// TIA Portal V21 export
ORGANIZATION_BLOCK "Pair"   // OB1, LAD
BEGIN

REGION Network 1: Motor
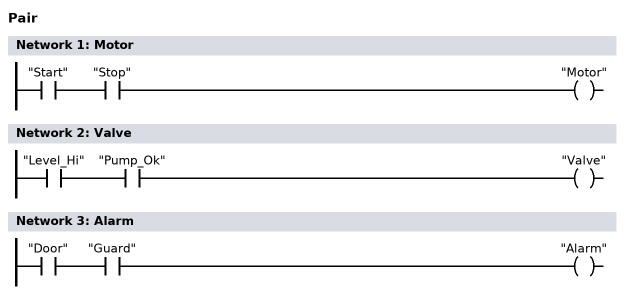
   RUNG wire#powerrail
      Contact( "Start" )
      Contact( "Stop" )
      Coil( "Motor" )
   END_RUNG
   // the same network as SCL:
   "Motor" := "Start" AND "Stop";
END_REGION

REGION Network 2: Valve
   RUNG wire#powerrail
      Contact( "Level_Hi" )
      Contact( "Pump_Ok" )
      Coil( "Valve" )
   END_RUNG
   // the same network as SCL:
   "Valve" := "Level_Hi" AND "Pump_Ok";
END_REGION

REGION Network 3: Alarm
   RUNG wire#powerrail
      Contact( "Door" )
      Contact( "Guard" )
      Coil( "Alarm" )
   END_RUNG
   // the same network as SCL:
   "Alarm" := "Door" AND "Guard";
END_REGION
END_ORGANIZATION_BLOCK
